// TIA Portal V20 export
DATA_BLOCK "T7_Datos"   // DB44900
{ S7_Optimized_Access := 'TRUE' }
AUTHOR : IA
FAMILY : PRUEBA
VERSION : 0.1
// Tanda 3: datos
// stored: AutoNumber false
   VAR
      Falso : Bool := false;
      Verdadero : Bool := true;
      Jmp_Fallo : Bool;
      Jmp_Llega : Bool;
      Jmpn_Fallo : Bool;
      Jmpn_Llega : Bool;
      UInt_1 : UInt := 1;
      JL_Fallo : Bool;
      JL_Llega : Bool;
      Int_5 : Int := 5;
      Int_3 : Int := 3;
      SW_Fallo : Bool;
      SW_Llega : Bool;
      Int_10 : Int := 10;
      VarGet_Out : Int;
      VarPut_Dst : Int;
      Int_7 : Int := 7;
      DInt_3 : DInt := 3;
      Int_42 : Int := 42;
      Ret_Write : Int := -1;
      Ret_Read : Int := -1;
      ArrDB_Leido : Int;
      Ret_Attr : Int := -1;
      DB_Longitud : UDInt;
      DB_Atributos : Byte;
      Ret_DIS_AIRT : Int := -1;
      Ret_EN_AIRT : Int := -1;
      SrtDint_Mem : Bool;
      Ret_SRT_DINT : Int := -1;
      T_100ms : Time := T#100MS;
      Word_0 : Word := 16#0;
      OB20_Cuenta : DInt;   // Lo incrementa el OB20 (alarma de retardo)
      Ret_QRY_DINT : Int := -1;
      St_QRY_DINT : Word;
      Ret_QRY_CINT : Int := -1;
      Ciclo_OB30 : UDInt;
      Fase_OB30 : UDInt;
      St_QRY_CINT : Word;
      OB30_Cuenta : DInt;   // Lo incrementa el OB30 (alarma cíclica)
      Ret_RTM : Int := -1;
      RTM_CQ : Bool;
      RTM_CV : DInt;
      Byte_0 : Byte := 16#0;
      DInt_0 : DInt := 0;
      Tog : Bool;
   END_VAR
BEGIN
END_DATA_BLOCK
